(* IEC 61131-3 sources: Gen-AI/final/Gen-AI_v1.0_submission/A2_框架源码/agent/logs/full34_fixture/E3_S06_1_42, 3 files *)

(* ---- best.st ---- *)
FUNCTION_BLOCK FB_S06
VAR_INPUT
    TempPV : REAL;
    SetTemp : REAL;
    Segment : INT;
    LoadReduceReq : BOOL;
END_VAR
VAR_OUTPUT
    HeatOn : BOOL;
    FanOn : BOOL;
    OverTempAlarm : BOOL;
    LoadReduce : BOOL;
    Status : WORD;
END_VAR
(* Add a VAR block for internal state/timers before the implementation, if needed. *)
(* SKELETON ONLY: replace this RETURN with scan logic and required initial state. *)
RETURN;
END_FUNCTION_BLOCK

(*  *)

(* ---- final.st ---- *)
FUNCTION_BLOCK FB_S06
VAR_INPUT
    TempPV : REAL;
    SetTemp : REAL;
    Segment : INT;
    LoadReduceReq : BOOL;
END_VAR
VAR_OUTPUT
    HeatOn : BOOL;
    FanOn : BOOL;
    OverTempAlarm : BOOL;
    LoadReduce : BOOL;
    Status : WORD;
END_VAR
(* Add a VAR block for internal state/timers before the implementation, if needed. *)
(* SKELETON ONLY: replace this RETURN with scan logic and required initial state. *)
RETURN;
END_FUNCTION_BLOCK

(*  *)

(* ---- skeleton.st ---- *)
FUNCTION_BLOCK FB_S06
VAR_INPUT
    TempPV : REAL;
    SetTemp : REAL;
    Segment : INT;
    LoadReduceReq : BOOL;
END_VAR
VAR_OUTPUT
    HeatOn : BOOL;
    FanOn : BOOL;
    OverTempAlarm : BOOL;
    LoadReduce : BOOL;
    Status : WORD;
END_VAR
(* Add a VAR block for internal state/timers before the implementation, if needed. *)
(* SKELETON ONLY: replace this RETURN with scan logic and required initial state. *)
RETURN;
END_FUNCTION_BLOCK
